Fanuc KAREL source: kt00568.KL

-- PROVISIONAL review KL for V940-1; original PC SHA256 a3c642527c1dd13d3f3f1e61dd814efeb631595cb7c3c113e7a9cb9278e28b72
-- Incomplete behavior may be omitted. Consult companion uncertainty JSON. Do not deploy.
PROGRAM KT00568
%NOLOCKGROUP
VAR
  R2 : REAL
-- UNRESOLVED_DECL V1 type=000013
-- UNRESOLVED_DECL OUT type=000013
BEGIN
  -- V9_ZERO_TABLE_METADATA_HINT layout=0001; no indexed target words; source/name/runtime held
  -- UNRESOLVED_PC offsets 5-20; opcodes 2E,22,32,35
  -- UNRESOLVED_PC offsets 25-36; opcodes 2E,23
  -- UNRESOLVED_PC offsets 41-63; opcodes 49,21,8E,4A
  -- UNRESOLVED_PC offsets 68-72; opcodes 7F
END KT00568
